Fanuc KAREL source: kx00013.KL

-- PROVISIONAL review KL for V1013-1; original PC SHA256 e930daa3e563ab9b345ddcd8df48857f0357e935baace56393e930e550cbefc9
-- Incomplete behavior may be omitted. Consult companion uncertainty JSON. Do not deploy.
PROGRAM KX00013
%NOLOCKGROUP
VAR
  I : INTEGER
  J : INTEGER
  B : BOOLEAN
  F : FILE
  S : STRING[80]
-- UNRESOLVED_DECL P type=000102
BEGIN
  -- UNRESOLVED_PC offsets 5-7; opcodes 9C,4E
  -- UNRESOLVED_PC offsets 12-16; opcodes 7F
END KX00013
